(* IEC 61131-3 sources: ArdisCVDCore/codesys, 27 files *)

(* ---- E_GasChannelInit.st ---- *)
TYPE E_GasChannelInit :
(
    INIT_START,
    INIT_RAMPTIME_HOLD,
    INIT_RAMPSTEP_HOLD,
    INIT_RAMPEN_HOLD,
    INIT_MODE_HOLD,
    INIT_DONE,
    CLOSE_HOLD,
    CLOSED
);
END_TYPE

(* ---- E_MicrowaveState.st ---- *)
TYPE E_MicrowaveState :
(
    MW_IDLE,
    MW_PREHEAT_START_HOLD,
    MW_PREHEATING,
    MW_PREHEAT_READY,
    MW_RUN_START_HOLD,
    MW_RUNNING,
    MW_RUN_STOP_HOLD,
    MW_PREHEAT_ABORT_HOLD,
    MW_FAULT_STOP_HOLD,
    MW_FAULT_LATCHED
);
END_TYPE

(* ---- ST_GasChannelState.st ---- *)
TYPE ST_GasChannelState :
STRUCT
    eInit            : E_GasChannelInit;
    iInitDelay       : INT;
    xRegulating      : BOOL;
    xFaultActive     : BOOL;
    xCloseConfirmed  : BOOL;
    iLastSetpointRaw : INT;
END_STRUCT
END_TYPE

(* ---- ST_MicrowaveState.st ---- *)
TYPE ST_MicrowaveState :
STRUCT
    xLastPreheatValue    : BOOL;
    xLastOnValue         : BOOL;
    xLastResetRequest    : BOOL;
    iLastSetpointRaw     : INT;
    wFaultReason         : WORD;
    iResetHoldScans      : INT;
    iPreheatElapsedScans : INT;
END_STRUCT
END_TYPE

(* ---- GVL_Alarms.st ---- *)
VAR_GLOBAL RETAIN
    wRetainMagic      : WORD;
    wParamAlarmEnable : WORD;
    wParamAbortEnable : WORD;
    abParamAlarmPct   : ARRAY[0..6] OF BYTE;
    abParamAbortPct   : ARRAY[0..6] OF BYTE;
    wMwReflAlarmWatt  : WORD;
    wMwReflAbortWatt  : WORD;
    wTempEnable       : WORD;
    wSampleTargetC    : WORD;
    bSampleAlarmPct   : BYTE;
    abWaterTargetC    : ARRAY[0..3] OF BYTE;
    abWaterAlarmPct   : ARRAY[0..3] OF BYTE;
    abWaterAbortPct   : ARRAY[0..3] OF BYTE;
    wInputEnable      : WORD;
    wInputReaction    : WORD;
    uiLidInput        : UINT;
END_VAR

VAR_GLOBAL
    awAlarmMask     : ARRAY[0..3] OF WORD;
    awAbortMask     : ARRAY[0..3] OF WORD;
    awAbortLatched  : ARRAY[0..3] OF WORD;
    xAbortActive    : BOOL;
    xRunActive      : BOOL;
    wGpvInhibit     : WORD;
    wVpvInhibit     : WORD;
    xForeVacInhibit : BOOL;
    xTurboInhibit   : BOOL;
    xMwInhibit      : BOOL;
    xMwTripActive   : BOOL;
    wMwTripLatched  : WORD;
    xThresholdsOk   : BOOL;
    xRetainWasBlank : BOOL;
    uiAbortCount    : UINT;
END_VAR

(* ---- GVL_CoolingIO.st ---- *)
VAR_GLOBAL
    awCoolMod1Value  : ARRAY[0..7] OF WORD;
    awCoolMod1Status : ARRAY[0..7] OF WORD;

    awCoolMod2Value  : ARRAY[0..7] OF WORD;
    awCoolMod2Status : ARRAY[0..7] OF WORD;
END_VAR

(* ---- GVL_Debug.st ---- *)
VAR_GLOBAL
    uiDbgGasReinitCount : UINT;
    xDbgReboot          : BOOL;
END_VAR

(* ---- GVL_GasIO.st ---- *)
VAR_GLOBAL
    awMeasuredRaw     : ARRAY[0..5] OF WORD;
    awSetpointRaw     : ARRAY[0..5] OF WORD;
    axSetpointTrigger : ARRAY[0..5] OF BOOL;

    awModeValue       : ARRAY[0..5] OF WORD;
    axModeTrigger     : ARRAY[0..5] OF BOOL;

    awRampTimeValue   : ARRAY[0..5] OF WORD;
    axRampTimeTrigger : ARRAY[0..5] OF BOOL;

    awRampStepValue   : ARRAY[0..5] OF WORD;
    axRampStepTrigger : ARRAY[0..5] OF BOOL;

    awRampEnValue     : ARRAY[0..5] OF WORD;
    axRampEnTrigger   : ARRAY[0..5] OF BOOL;
END_VAR

(* ---- GVL_GasValveIO.st ---- *)
VAR_GLOBAL
    axGpvOutput : ARRAY[1..8] OF BOOL;
END_VAR

(* ---- GVL_MicrowaveIO.st ---- *)
VAR_GLOBAL
    awMwPowerRaw       : ARRAY[0..1] OF WORD;
    axMwStatusBlock1   : ARRAY[0..1] OF BOOL;
    axMwStatusBlock2   : ARRAY[0..5] OF BOOL;
    axMwStatusBlock3   : ARRAY[0..7] OF BOOL;

    xMwPreheatValue    : BOOL;
    xMwPreheatTrigger  : BOOL;
    xMwOnValue         : BOOL;
    xMwOnTrigger       : BOOL;
    xMwResetTrigger    : BOOL;
    wMwSetpointRaw     : WORD;
    xMwSetpointTrigger : BOOL;
END_VAR

(* ---- GVL_ModbusHolding.st ---- *)
VAR_GLOBAL
    awHolding AT %QW0 : ARRAY[0..295] OF WORD;
END_VAR

(* ---- GVL_PlcIO.st ---- *)
VAR_GLOBAL
    axFastDigitalIn : ARRAY[1..8] OF BOOL;
    axDigitalIn     : ARRAY[9..12] OF BOOL;
END_VAR

(* ---- GVL_PyroIO.st ---- *)
VAR_GLOBAL
    awPyroRxtCh1Raw     : ARRAY[0..1] OF WORD;
    awPyroRxtCh2Raw     : ARRAY[0..1] OF WORD;
    awPyroRxtRatioRaw   : ARRAY[0..1] OF WORD;
    wPyroRxtAdcStatus   : WORD;
    wPyroRxtDevStatus   : WORD;

    awPyroSmartCh1Raw   : ARRAY[0..1] OF WORD;
    awPyroSmartCh2Raw   : ARRAY[0..1] OF WORD;
    awPyroSmartRatioRaw : ARRAY[0..1] OF WORD;
    wPyroSmartAdcStatus : WORD;
    wPyroSmartDevStatus : WORD;
END_VAR

(* ---- GVL_TurboPumpIO.st ---- *)
VAR_GLOBAL
    awTurboStatusRaw  : ARRAY[0..3] OF WORD;
    wTurboTempRaw     : WORD;

    wTurboCommandValue   : WORD;
    xTurboCommandTrigger : BOOL;
END_VAR

(* ---- GVL_VacuumIO.st ---- *)
VAR_GLOBAL
    axVpvOutput : ARRAY[1..8] OF BOOL;
    xWaterPumpOutput : BOOL;
    xForeVacPumpOutput : BOOL;
END_VAR

(* ---- FB_IncrementalPid.st ---- *)
FUNCTION_BLOCK FB_IncrementalPid
VAR_INPUT
    xEnable       : BOOL;
    xReset        : BOOL;
    xDirectMode   : BOOL;
    rSetpoint     : REAL;
    rMeasured     : REAL;
    rKp           : REAL;
    rKi           : REAL;
    rKd           : REAL;
    xSmartMode    : BOOL;
    rSmartKp      : REAL;
    wPresetId     : WORD;
    rPresetOutput : REAL;
    wShiftId      : WORD;
    rShiftDelta   : REAL;
    rLowerLimit   : REAL;
    rUpperLimit   : REAL;
    rDirectValue  : REAL;
    rCycleSeconds : REAL := 0.2;
END_VAR
VAR_OUTPUT
    rError  : REAL;
    rP      : REAL;
    rI      : REAL;
    rD      : REAL;
    rOutput : REAL;
    wPresetDoneId : WORD;
    wShiftDoneId  : WORD;
END_VAR
VAR
    rPreviousError : REAL;
    xInitialized   : BOOL;
    rMin           : REAL;
    rMax           : REAL;
	arErrorBuffer      : ARRAY[0..99] OF REAL;
    i                  : INT;
    rErrAverageFirst   : REAL;
    rErrAverageLast    : REAL;
    rErrAverageIntegral : REAL;
    rKpActive           : REAL;
    wPresetSeenId       : WORD;
    xPresetArmed        : BOOL;
    rPresetFromError    : REAL;
    wShiftSeenId        : WORD;
    xShiftNew           : BOOL;
    rPresetShift        : REAL;
END_VAR

IF rLowerLimit <= rUpperLimit THEN
    rMin := rLowerLimit;
    rMax := rUpperLimit;
ELSE
    rMin := rUpperLimit;
    rMax := rLowerLimit;
END_IF;

rError := rMeasured - rSetpoint;

xShiftNew := FALSE;
IF wShiftId <> wShiftSeenId THEN
    wShiftSeenId := wShiftId;
    IF wShiftId <> WORD#0 THEN
        xShiftNew := TRUE;
        wShiftDoneId := wShiftId;
    END_IF;
END_IF;

IF NOT xEnable THEN
    rP := 0.0;
    rI := 0.0;
    rD := 0.0;
    rOutput := rMin;
    rPreviousError := rError;
    xInitialized := FALSE;
    RETURN;
END_IF;

IF xReset OR NOT xInitialized THEN
    rPreviousError := rError;
    rOutput := rMin;

    FOR i := 0 TO 99 DO
        arErrorBuffer[i] := rError;
    END_FOR;

    xInitialized := TRUE;
END_IF;

IF xShiftNew THEN
    IF xPresetArmed THEN
        rPresetShift := rPresetShift + rShiftDelta;
    ELSIF NOT xDirectMode THEN
        rOutput := rOutput + rShiftDelta;
    END_IF;
END_IF;

IF wPresetId <> wPresetSeenId THEN
    wPresetSeenId := wPresetId;
    xPresetArmed := wPresetId <> WORD#0;
    rPresetFromError := rError;
    rPresetShift := 0.0;
END_IF;

IF rCycleSeconds > 0.001 THEN
    FOR i := 0 TO 98 DO
        arErrorBuffer[i] := arErrorBuffer[i + 1];
    END_FOR;
    arErrorBuffer[99] := rError;

    rErrAverageFirst := 0.0;
    FOR i := 87 TO 91 DO
        rErrAverageFirst := rErrAverageFirst + arErrorBuffer[i];
    END_FOR;
    rErrAverageFirst := rErrAverageFirst / 5.0;

    rErrAverageLast := 0.0;
    FOR i := 98 TO 99 DO
        rErrAverageLast := rErrAverageLast + arErrorBuffer[i];
    END_FOR;
    rErrAverageLast := rErrAverageLast / 2.0;

    rD := rKd * (rErrAverageLast - rErrAverageFirst);

    rErrAverageIntegral := 0.0;
    FOR i := 80 TO 99 DO
        rErrAverageIntegral := rErrAverageIntegral + arErrorBuffer[i];
    END_FOR;
    rErrAverageIntegral := rErrAverageIntegral / 20.0;

    rI := rKi * rErrAverageIntegral;
ELSE
    rD := 0.0;
    rI := 0.0;
END_IF;

IF xSmartMode AND rError > 0.0 AND rD > 0.0 THEN
    rKpActive := rSmartKp;
ELSE
    rKpActive := rKp;
END_IF;

rP := rKpActive * rError;

rPreviousError := rError;

IF xDirectMode THEN
    rOutput := rDirectValue;
    rPresetFromError := rError;
ELSIF xPresetArmed AND rError * rPresetFromError <= 0.0 THEN
    rOutput := rPresetOutput + rPresetShift;
    xPresetArmed := FALSE;
    wPresetDoneId := wPresetSeenId;
ELSE
    rOutput := rOutput + rP + rI + rD;
END_IF;

IF rOutput > rMax THEN
    rOutput := rMax;
ELSIF rOutput < rMin THEN
    rOutput := rMin;
END_IF;

(* ---- FB_ThyracontAscii.st ---- *)
FUNCTION_BLOCK FB_ThyracontAscii
VAR_INPUT
    xEnable : BOOL := TRUE;
    udiPort : UDINT := 1;
    udiAddress : UDINT := 1;
    udiBaudrate : UDINT := 9600;
    tPollInterval : TIME := T#1S;
END_VAR
VAR_OUTPUT
    xValid : BOOL;
    xConnected : BOOL;
    rPressureMbar : REAL;
    rPressureTorr : REAL;
    wStatusFlags : WORD;
    wErrorCode : WORD;
    udiCycle : UDINT;
END_VAR
VAR
    fbOpen : COM.Open;
    fbWrite : COM.Write;
    fbRead : COM.Read;
    aParams : ARRAY[1..7] OF COM.PARAMETER;
    hCom : CAA.HANDLE;
    aTx : ARRAY[0..9] OF BYTE := [BYTE#48, BYTE#48, BYTE#49, BYTE#48, BYTE#77, BYTE#86, BYTE#48, BYTE#48, BYTE#68, BYTE#13];
    aRx : ARRAY[0..63] OF BYTE;
    aAdr : ARRAY[0..2] OF BYTE;
    iAddr : INT;
    iChecksum : INT;
    iState : INT;
    udiPollTicks : UDINT;
    udiPollTicksMax : UDINT := 5;
    xOpenExecute : BOOL;
    xWriteExecute : BOOL;
    xReadExecute : BOOL;
    i : INT;
    j : INT;
    iSize : INT;
    iFrameStart : INT;
    iDataLen : INT;
    iDataStart : INT;
    iDigit : INT;
    iSign : INT;
    iExpSign : INT;
    iExp : INT;
    rParsed : REAL;
    rDiv : REAL;
    xFraction : BOOL;
    xExponent : BOOL;
    xHasDigit : BOOL;
END_VAR

IF NOT xEnable THEN
    xOpenExecute := FALSE;
    xWriteExecute := FALSE;
    xReadExecute := FALSE;
    xConnected := FALSE;
    xValid := FALSE;
    wStatusFlags := WORD#0;
    wErrorCode := WORD#0;
    iState := 0;
    RETURN;
END_IF;

aParams[1].udiParameterId := COM.CAA_Parameter_Constants.udiPort;
aParams[1].udiValue := udiPort;
aParams[2].udiParameterId := COM.CAA_Parameter_Constants.udiBaudrate;
aParams[2].udiValue := udiBaudrate;
aParams[3].udiParameterId := COM.CAA_Parameter_Constants.udiParity;
aParams[3].udiValue := 2;
aParams[4].udiParameterId := COM.CAA_Parameter_Constants.udiStopBits;
aParams[4].udiValue := 0;
aParams[5].udiParameterId := COM.CAA_Parameter_Constants.udiTimeout;
aParams[5].udiValue := 200000;
aParams[6].udiParameterId := COM.CAA_Parameter_Constants.udiByteSize;
aParams[6].udiValue := 8;
aParams[7].udiParameterId := COM.CAA_Parameter_Constants.udiBinary;
aParams[7].udiValue := 1;

iAddr := UDINT_TO_INT(udiAddress);
IF (iAddr < 1) OR (iAddr > 16) THEN
    iAddr := 1;
END_IF;
aAdr[0] := INT_TO_BYTE(iAddr / 100 MOD 10 + 48);
aAdr[1] := INT_TO_BYTE(iAddr / 10 MOD 10 + 48);
aAdr[2] := INT_TO_BYTE(iAddr MOD 10 + 48);
aTx[0] := aAdr[0];
aTx[1] := aAdr[1];
aTx[2] := aAdr[2];

iChecksum := 0;
FOR i := 0 TO 7 DO
    iChecksum := iChecksum + BYTE_TO_INT(aTx[i]);
END_FOR;
aTx[8] := INT_TO_BYTE(iChecksum MOD 64 + 64);

IF tPollInterval <= T#0MS THEN
    udiPollTicksMax := 0;
ELSIF tPollInterval <= T#200MS THEN
    udiPollTicksMax := 1;
ELSE
    udiPollTicksMax := TIME_TO_UDINT(tPollInterval) / 200;
    IF udiPollTicksMax < 1 THEN
        udiPollTicksMax := 1;
    END_IF;
END_IF;

CASE iState OF
    0:
        xOpenExecute := TRUE;
        xConnected := FALSE;
        xValid := FALSE;
        wErrorCode := WORD#1;
        IF fbOpen.xDone THEN
            hCom := fbOpen.hCom;
            xOpenExecute := FALSE;
            xConnected := TRUE;
            wErrorCode := WORD#0;
            iState := 10;
        ELSIF fbOpen.xError THEN
            xOpenExecute := FALSE;
            wErrorCode := WORD#2;
            iState := 50;
        END_IF;

    10:
        udiPollTicks := 0;
        FOR i := 0 TO 63 DO
            aRx[i] := BYTE#0;
        END_FOR;
        xWriteExecute := TRUE;
        iState := 20;

    20:
        IF fbWrite.xDone THEN
            xWriteExecute := FALSE;
            xReadExecute := TRUE;
            iState := 30;
        ELSIF fbWrite.xError THEN
            xWriteExecute := FALSE;
            xValid := FALSE;
            wErrorCode := WORD#3;
            iState := 50;
        END_IF;

    30:
        IF fbRead.xDone THEN
            xReadExecute := FALSE;
            iSize := UDINT_TO_INT(fbRead.szSize);
            iFrameStart := -1;

            IF iSize >= 10 THEN
                FOR i := 0 TO iSize - 8 DO
                    IF (aRx[i] = aAdr[0]) AND (aRx[i + 1] = aAdr[1]) AND
                       (aRx[i + 2] = aAdr[2]) AND (aRx[i + 3] = BYTE#49) AND
                       (aRx[i + 4] = BYTE#77) AND (aRx[i + 5] = BYTE#86) THEN
                        iFrameStart := i;
                        EXIT;
                    END_IF;
                END_FOR;
            END_IF;

            IF iFrameStart < 0 THEN
                xValid := FALSE;
                wErrorCode := WORD#5;
                iState := 50;
            ELSE
                iDataLen := (BYTE_TO_INT(aRx[iFrameStart + 6]) - 48) * 10 +
                            (BYTE_TO_INT(aRx[iFrameStart + 7]) - 48);
                iDataStart := iFrameStart + 8;

                IF (iDataLen <= 0) OR ((iDataStart + iDataLen) >= iSize) THEN
                    xValid := FALSE;
                    wErrorCode := WORD#6;
                    iState := 50;
                ELSE
                    rParsed := 0.0;
                    rDiv := 10.0;
                    iSign := 1;
                    iExpSign := 1;
                    iExp := 0;
                    xFraction := FALSE;
                    xExponent := FALSE;
                    xHasDigit := FALSE;

                    FOR i := 0 TO iDataLen - 1 DO
                        j := iDataStart + i;
                        IF (aRx[j] >= BYTE#48) AND (aRx[j] <= BYTE#57) THEN
                            iDigit := BYTE_TO_INT(aRx[j]) - 48;
                            xHasDigit := TRUE;
                            IF xExponent THEN
                                iExp := iExp * 10 + iDigit;
                            ELSIF xFraction THEN
                                rParsed := rParsed + INT_TO_REAL(iDigit) / rDiv;
                                rDiv := rDiv * 10.0;
                            ELSE
                                rParsed := rParsed * 10.0 + INT_TO_REAL(iDigit);
                            END_IF;
                        ELSIF aRx[j] = BYTE#45 THEN
                            IF xExponent THEN
                                iExpSign := -1;
                            ELSE
                                iSign := -1;
                            END_IF;
                        ELSIF (aRx[j] = BYTE#46) OR (aRx[j] = BYTE#44) THEN
                            xFraction := TRUE;
                        ELSIF (aRx[j] = BYTE#69) OR (aRx[j] = BYTE#101) THEN
                            xExponent := TRUE;
                        END_IF;
                    END_FOR;

                    IF xHasDigit THEN
                        IF iExp > 38 THEN
                            iExp := 38;
                        END_IF;

                        FOR i := 1 TO iExp DO
                            IF iExpSign > 0 THEN
                                rParsed := rParsed * 10.0;
                            ELSE
                                rParsed := rParsed / 10.0;
                            END_IF;
                        END_FOR;

                        rPressureMbar := rParsed * INT_TO_REAL(iSign);
                        rPressureTorr := rPressureMbar * 0.7500637;
                        xValid := TRUE;
                        xConnected := TRUE;
                        wErrorCode := WORD#0;
                        udiCycle := udiCycle + 1;
                    ELSE
                        xValid := FALSE;
                        wErrorCode := WORD#7;
                    END_IF;

                    iState := 50;
                END_IF;
            END_IF;
        ELSIF fbRead.xError THEN
            xReadExecute := FALSE;
            xValid := FALSE;
            wErrorCode := WORD#4;
            iState := 50;
        END_IF;

    50:
        udiPollTicks := udiPollTicks + 1;
        IF udiPollTicks >= udiPollTicksMax THEN
            iState := 10;
        END_IF;

ELSE
    iState := 0;
END_CASE;

wStatusFlags := WORD#0;
IF xValid THEN
    wStatusFlags := wStatusFlags OR WORD#16#0001;
END_IF;

fbOpen(
    xExecute := xOpenExecute,
    usiListLength := 7,
    pParameterList := ADR(aParams));

fbWrite(
    xExecute := xWriteExecute,
    udiTimeOut := 100000,
    hCom := hCom,
    pBuffer := ADR(aTx),
    szSize := SIZEOF(aTx));

fbRead(
    xExecute := xReadExecute,
    udiTimeOut := 300000,
    hCom := hCom,
    pBuffer := ADR(aRx),
    szBuffer := SIZEOF(aRx));

(* ---- PLC_PRG.st ---- *)
PROGRAM PLC_PRG
(* main program: hmi link, signal tower, pressure pid *)
VAR
    xDoBlinkTest : BOOL;
    wBenchMuAo1Output : ARRAY[0..0] OF WORD;
    xTrafficLightGreen  : BOOL;
    xTrafficLightYellow : BOOL;
    xTrafficLightRed    : BOOL;
    wTrafficLightMask   : WORD;

    xHmiWriteSeen         : BOOL;
    udiHmiStaleCycles     : UDINT;
    xHmiLinkLost          : BOOL;

    awMvAi1Value  : ARRAY[0..1] OF WORD;
    awMvAi1Status : ARRAY[0..0] OF WORD;
    uMvAi1Value   : U_DWORD_REAL;
    wMvAi1Status  : WORD;
    xMvAi1Ok      : BOOL;
    rMvAi1Percent : REAL;
    rMvAi1Voltage : REAL;
    rChMeasuredMv : REAL;

	wDiscreteInputs : WORD;
    iDiIndex        : INT;

    rChamberMuAo1Command : REAL;
    xChamberMuAo1Clamped : BOOL;
    uiChamberMuAo1Command : UINT;
    fbChamber : FB_IncrementalPid;
    fbPlenum  : FB_IncrementalPid;
    xProtocolOk    : BOOL;
    xChamberEnable : BOOL;
    xPlenumEnable  : BOOL;
    xReset         : BOOL;
    udiCycle       : UDINT;
    rChSetpoint : REAL;
    rChMeasured : REAL;
    rChKp       : REAL;
    rChKi       : REAL;
    rChKd       : REAL;
    rChLower    : REAL;
    rChUpper    : REAL;
    rChDirect   : REAL;
    rChSmartKp  : REAL;
    xChSmartMode : BOOL;
    rChPresetOutput : REAL;
    wChPresetId     : WORD;
    rChShiftDelta   : REAL;
    wChShiftId      : WORD;
    rPlSetpoint : REAL;
    rPlMeasured : REAL;
    rPlKp       : REAL;
    rPlKi       : REAL;
    rPlKd       : REAL;
    rPlLower    : REAL;
    rPlUpper    : REAL;
    rPlDirect   : REAL;
    dwValue     : DWORD;
    xDoBlinkTestEnable : BOOL;
    xBenchMuAo1Enable : BOOL;
    xBenchMuAo1Clamped : BOOL;
    uiBenchMuAo1Command : UINT;
    uiBenchMuAo1Applied : UINT;
    awMvAi1Raw : ARRAY[0..1] OF WORD;
END_VAR
VAR CONSTANT
    HMI_STALE_CYCLES  : UDINT := UDINT#15;
END_VAR

(* commands from the hmi *)
xProtocolOk := awHolding[0] = WORD#1;
xChamberEnable := xProtocolOk AND (awHolding[1] AND WORD#16#0001) <> WORD#0;
xPlenumEnable := xProtocolOk AND (awHolding[1] AND WORD#16#0002) <> WORD#0;
xReset := (awHolding[1] AND WORD#16#0004) <> WORD#0;
xTrafficLightGreen  := (awHolding[1] AND WORD#16#0010) <> WORD#0;
xTrafficLightYellow := (awHolding[1] AND WORD#16#0020) <> WORD#0;
xTrafficLightRed    := (awHolding[1] AND WORD#16#0040) <> WORD#0;

(* hmi watchdog: link lost after 3 s without a write *)
xHmiWriteSeen := (awHolding[1] AND WORD#16#8000) = WORD#0;

IF xHmiWriteSeen THEN
    udiHmiStaleCycles := UDINT#0;
ELSIF udiHmiStaleCycles < HMI_STALE_CYCLES THEN
    udiHmiStaleCycles := udiHmiStaleCycles + UDINT#1;
END_IF;

xHmiLinkLost := udiHmiStaleCycles >= HMI_STALE_CYCLES;

(* signal tower, all three lamps on when the link is lost *)
wTrafficLightMask := WORD#0;
IF xHmiLinkLost THEN
    wTrafficLightMask := WORD#16#0007;
ELSE
    IF xTrafficLightGreen THEN
        wTrafficLightMask := wTrafficLightMask OR WORD#16#0001;
    END_IF;
    IF xTrafficLightYellow THEN
        wTrafficLightMask := wTrafficLightMask OR WORD#16#0002;
    END_IF;
    IF xTrafficLightRed THEN
        wTrafficLightMask := wTrafficLightMask OR WORD#16#0004;
    END_IF;
END_IF;

(* set the marker, the hmi clears it on its next write *)
awHolding[1] := awHolding[1] OR WORD#16#8000;

(* chamber pid output to the analogue output, max 500 *)
rChamberMuAo1Command := fbChamber.rOutput / 10.0;
xChamberMuAo1Clamped := rChamberMuAo1Command > 500.0;

IF xChamberMuAo1Clamped THEN
    uiChamberMuAo1Command := UINT#500;
ELSE
    uiChamberMuAo1Command := REAL_TO_UINT(rChamberMuAo1Command);
END_IF;

(* chamber pressure from the analogue input module *)
wMvAi1Status := awMvAi1Status[0];
xMvAi1Ok := wMvAi1Status = WORD#16#0000;

uMvAi1Value.dwValue := SHL(WORD_TO_DWORD(awMvAi1Value[1]), 16) OR WORD_TO_DWORD(awMvAi1Value[0]);
rMvAi1Percent := uMvAi1Value.rValue;
rMvAi1Voltage := LIMIT(0.0, rMvAi1Percent / 10.0, 10.0);

IF xMvAi1Ok THEN
    rChMeasuredMv := LIMIT(0.0, rMvAi1Percent * 10.0, 1000.0);
END_IF;

(* pid setpoints and gains from the hmi *)
rChSetpoint := F_ReadFixed(awHolding[4], awHolding[5]);
rChMeasured := rChMeasuredMv;
rChKp := F_ReadFixed(awHolding[8], awHolding[9]);
rChKi := F_ReadFixed(awHolding[10], awHolding[11]);
rChKd := F_ReadFixed(awHolding[12], awHolding[13]);
rChLower := F_ReadFixed(awHolding[14], awHolding[15]);
rChUpper := F_ReadFixed(awHolding[16], awHolding[17]);
rChDirect := F_ReadFixed(awHolding[18], awHolding[19]);
rChSmartKp := F_ReadFixed(awHolding[27], awHolding[28]);
xChSmartMode := awHolding[29] <> WORD#0;
rChPresetOutput := F_ReadFixed(awHolding[56], awHolding[57]);
wChPresetId := awHolding[58];
rChShiftDelta := F_ReadFixed(awHolding[59], awHolding[60]);
wChShiftId := awHolding[61];

rPlSetpoint := F_ReadFixed(awHolding[30], awHolding[31]);
rPlMeasured := F_ReadFixed(awHolding[32], awHolding[33]);
rPlKp := F_ReadFixed(awHolding[34], awHolding[35]);
rPlKi := F_ReadFixed(awHolding[36], awHolding[37]);
rPlKd := F_ReadFixed(awHolding[38], awHolding[39]);
rPlLower := F_ReadFixed(awHolding[40], awHolding[41]);
rPlUpper := F_ReadFixed(awHolding[42], awHolding[43]);
rPlDirect := F_ReadFixed(awHolding[44], awHolding[45]);

(* chamber pid *)
fbChamber(
    xEnable := xChamberEnable,
    xReset := xReset,
    xDirectMode := awHolding[20] <> WORD#0,
    rSetpoint := rChSetpoint,
    rMeasured := rChMeasured,
    rKp := rChKp,
    rKi := rChKi,
    rKd := rChKd,
    xSmartMode := xChSmartMode,
    rSmartKp := rChSmartKp,
    wPresetId := wChPresetId,
    rPresetOutput := rChPresetOutput,
    wShiftId := wChShiftId,
    rShiftDelta := rChShiftDelta,
    rLowerLimit := rChLower,
    rUpperLimit := rChUpper,
    rDirectValue := rChDirect,
    rCycleSeconds := 0.2);

(* plenum pid *)
fbPlenum(
    xEnable := xPlenumEnable,
    xReset := xReset,
    xDirectMode := awHolding[46] <> WORD#0,
    rSetpoint := rPlSetpoint,
    rMeasured := rPlMeasured,
    rKp := rPlKp,
    rKi := rPlKi,
    rKd := rPlKd,
    rLowerLimit := rPlLower,
    rUpperLimit := rPlUpper,
    rDirectValue := rPlDirect,
    rCycleSeconds := 0.2);

(* cycle counter and blink test *)
udiCycle := udiCycle + 1;
xDoBlinkTestEnable := awHolding[150] = WORD#16#A55A;
xDoBlinkTest := xDoBlinkTestEnable AND ((udiCycle MOD UDINT#10) < UDINT#5);

(* to the hmi: version, status, cycle counter *)
awHolding[100] := WORD#1;
IF xProtocolOk THEN
    awHolding[101] := WORD#16#0003;
ELSE
    awHolding[101] := WORD#0;
END_IF;
awHolding[102] := DWORD_TO_WORD(udiCycle);
awHolding[103] := DWORD_TO_WORD(SHR(udiCycle, 16));

(* chamber pid terms to the hmi *)
dwValue := F_ToFixed(fbChamber.rError);
awHolding[104] := DWORD_TO_WORD(dwValue);
awHolding[105] := DWORD_TO_WORD(SHR(dwValue, 16));
dwValue := F_ToFixed(fbChamber.rP);
awHolding[106] := DWORD_TO_WORD(dwValue);
awHolding[107] := DWORD_TO_WORD(SHR(dwValue, 16));
dwValue := F_ToFixed(fbChamber.rI);
awHolding[108] := DWORD_TO_WORD(dwValue);
awHolding[109] := DWORD_TO_WORD(SHR(dwValue, 16));
dwValue := F_ToFixed(fbChamber.rD);
awHolding[110] := DWORD_TO_WORD(dwValue);
awHolding[111] := DWORD_TO_WORD(SHR(dwValue, 16));
dwValue := F_ToFixed(fbChamber.rOutput);
awHolding[112] := DWORD_TO_WORD(dwValue);
awHolding[113] := DWORD_TO_WORD(SHR(dwValue, 16));
awHolding[114] := fbChamber.wPresetDoneId;
awHolding[115] := fbChamber.wShiftDoneId;

(* plenum pid terms to the hmi *)
dwValue := F_ToFixed(fbPlenum.rError);
awHolding[120] := DWORD_TO_WORD(dwValue);
awHolding[121] := DWORD_TO_WORD(SHR(dwValue, 16));
dwValue := F_ToFixed(fbPlenum.rP);
awHolding[122] := DWORD_TO_WORD(dwValue);
awHolding[123] := DWORD_TO_WORD(SHR(dwValue, 16));
dwValue := F_ToFixed(fbPlenum.rI);
awHolding[124] := DWORD_TO_WORD(dwValue);
awHolding[125] := DWORD_TO_WORD(SHR(dwValue, 16));
dwValue := F_ToFixed(fbPlenum.rD);
awHolding[126] := DWORD_TO_WORD(dwValue);
awHolding[127] := DWORD_TO_WORD(SHR(dwValue, 16));
dwValue := F_ToFixed(fbPlenum.rOutput);
awHolding[128] := DWORD_TO_WORD(dwValue);
awHolding[129] := DWORD_TO_WORD(SHR(dwValue, 16));

(* chamber pressure and sensor status to the hmi *)
dwValue := F_ToFixed(rChMeasuredMv);
awHolding[130] := DWORD_TO_WORD(dwValue);
awHolding[131] := DWORD_TO_WORD(SHR(dwValue, 16));
awHolding[132] := wMvAi1Status;

(* discrete inputs to the hmi *)
wDiscreteInputs := WORD#0;
FOR iDiIndex := 1 TO 8 DO
    IF axFastDigitalIn[iDiIndex] THEN
        wDiscreteInputs := wDiscreteInputs OR SHL(WORD#1, iDiIndex - 1);
    END_IF;
END_FOR;
FOR iDiIndex := 9 TO 12 DO
    IF axDigitalIn[iDiIndex] THEN
        wDiscreteInputs := wDiscreteInputs OR SHL(WORD#1, iDiIndex - 1);
    END_IF;
END_FOR;
awHolding[139] := wDiscreteInputs;

(* manual analogue output test from the hmi *)
uiBenchMuAo1Command := WORD_TO_UINT(awHolding[154]);
xBenchMuAo1Enable := awHolding[155] = WORD#16#A55A;
xBenchMuAo1Clamped := uiBenchMuAo1Command > UINT#500;

IF xBenchMuAo1Clamped THEN
    uiBenchMuAo1Command := UINT#500;
END_IF;

IF xBenchMuAo1Enable THEN
    uiBenchMuAo1Applied := uiBenchMuAo1Command;
ELSE
    uiBenchMuAo1Applied := UINT#0;
END_IF;

(* test flags to the hmi *)
IF xBenchMuAo1Enable THEN
    awHolding[157] := awHolding[157] OR WORD#16#0001;
END_IF;

IF xBenchMuAo1Clamped THEN
    awHolding[157] := awHolding[157] OR WORD#16#0002;
END_IF;

(* output command from the chamber pid *)
IF fbChamber.rOutput <= 0.0 THEN
    uiChamberMuAo1Command := UINT#0;
    xChamberMuAo1Clamped := FALSE;
ELSE
    rChamberMuAo1Command := fbChamber.rOutput / 10.0;
    xChamberMuAo1Clamped := rChamberMuAo1Command > 500.0;

    IF xChamberMuAo1Clamped THEN
        uiChamberMuAo1Command := UINT#500;
    ELSE
        uiChamberMuAo1Command := REAL_TO_UINT(rChamberMuAo1Command);
    END_IF;
END_IF;

(* drive the output: test value, pid or zero *)
IF xBenchMuAo1Enable THEN
    uiBenchMuAo1Applied := uiBenchMuAo1Command;
ELSIF xChamberEnable THEN
    uiBenchMuAo1Applied := uiChamberMuAo1Command;
ELSE
    uiBenchMuAo1Applied := UINT#0;
END_IF;

wBenchMuAo1Output[0] := UINT_TO_WORD(uiBenchMuAo1Applied);
awHolding[156] := wBenchMuAo1Output[0];

(* ---- PRG_Alarms.st ---- *)
PROGRAM PRG_Alarms
(* alarms and abort *)
VAR
    i : INT;
    iBase : INT;
    iBit : INT;
    iWord : INT;

    xFirstScan : BOOL := TRUE;

    axAlarm : ARRAY[0..63] OF BOOL;
    axAbort : ARRAY[0..63] OF BOOL;

    arBandSetpoint : ARRAY[0..6] OF REAL;
    arBandMeasured : ARRAY[0..6] OF REAL;
    axBandGate     : ARRAY[0..6] OF BOOL;

    arWaterTempC : ARRAY[0..3] OF REAL;
    axWaterTempValid : ARRAY[0..3] OF BOOL;

    rSetpoint : REAL;
    rMeasured : REAL;
    rBand     : REAL;
    rReflKw   : REAL;
    rSampleC  : REAL;
    rFlowLpm  : REAL;
    rWaterBar : REAL;
    rCdaBar   : REAL;

    wCommand    : WORD;
    wStatusWord : WORD;
    wMwStatus : WORD;
    wTempValid : WORD;
    wFlowValid : WORD;
    wTurboStatus : WORD;
    wDiscrete : WORD;
    wMwTripNow : WORD;

    xMwRequested : BOOL;
    xPyroValid : BOOL;
    xTurboAnswering : BOOL;
    xWaterPump : BOOL;
    xFlowArmed : BOOL;
    xLidClosed : BOOL;

    xAnyAlarm : BOOL;
    xAnyAbort : BOOL;

    xReset : BOOL;
    xResetPrev : BOOL;

    fbFlowArm : TON;
END_VAR
VAR CONSTANT
    C_BLOCK_MAGIC  : WORD := WORD#16#A500;
    C_RETAIN_MAGIC : WORD := WORD#16#5A5A;

    C_FLOW_MIN_LOW  : REAL := 1.0;
    C_FLOW_MIN_HIGH : REAL := 5.0;

    C_WATER_ALARM_BAR : REAL := 0.7;
    C_WATER_ABORT_BAR : REAL := 0.5;
    C_CDA_ALARM_BAR   : REAL := 5.0;
    C_CDA_ABORT_BAR   : REAL := 4.0;

    C_CHAMBER_MAX_TORR : REAL := 800.0;
    C_HMI_PROTOCOL     : WORD := WORD#16#0200;
    C_FLOW_ARM_TIME    : TIME := T#4S;

    C_CIRC_STAGE    : INT := 0;
    C_CIRC_CHAMBER  : INT := 1;
    C_CIRC_MWHEAD   : INT := 2;
    C_CIRC_MWPOWER  : INT := 3;
    C_CIRC_INTERNAL : INT := 5;
    C_CIRC_EXTERNAL : INT := 6;
END_VAR

(* first scan: all alarms off if the retain memory was lost *)
IF xFirstScan THEN
    xFirstScan := FALSE;
    IF wRetainMagic <> C_RETAIN_MAGIC THEN
        xRetainWasBlank := TRUE;
        wRetainMagic := C_RETAIN_MAGIC;
        wParamAlarmEnable := WORD#0;
        wParamAbortEnable := WORD#0;
        wTempEnable := WORD#0;
        wInputEnable := WORD#0;
        uiLidInput := UINT#1;
    ELSE
        xRetainWasBlank := FALSE;
    END_IF;
END_IF;

(* alarm thresholds from the hmi *)
xThresholdsOk := (awHolding[248] AND WORD#16#FF00) = C_BLOCK_MAGIC;

IF xThresholdsOk THEN
    wParamAlarmEnable := awHolding[249];
    wParamAbortEnable := awHolding[250];
    FOR i := 0 TO 6 DO
        abParamAlarmPct[i] := WORD_TO_BYTE(awHolding[251 + i] AND WORD#16#00FF);
        abParamAbortPct[i] := WORD_TO_BYTE(SHR(awHolding[251 + i], 8));
    END_FOR;
    wMwReflAlarmWatt := awHolding[258];
    wMwReflAbortWatt := awHolding[259];

    wTempEnable := awHolding[260];
    wSampleTargetC := awHolding[261];
    bSampleAlarmPct := WORD_TO_BYTE(awHolding[262] AND WORD#16#00FF);
    abWaterTargetC[0] := WORD_TO_BYTE(awHolding[263] AND WORD#16#00FF);
    abWaterTargetC[1] := WORD_TO_BYTE(SHR(awHolding[263], 8));
    abWaterTargetC[2] := WORD_TO_BYTE(awHolding[264] AND WORD#16#00FF);
    abWaterTargetC[3] := WORD_TO_BYTE(SHR(awHolding[264], 8));
    FOR i := 0 TO 3 DO
        abWaterAlarmPct[i] := WORD_TO_BYTE(awHolding[265 + i] AND WORD#16#00FF);
        abWaterAbortPct[i] := WORD_TO_BYTE(SHR(awHolding[265 + i], 8));
    END_FOR;

    wInputEnable := awHolding[269];
    wInputReaction := awHolding[270];
    xRunActive := (awHolding[271] AND WORD#16#0001) <> WORD#0;
    uiLidInput := WORD_TO_UINT(SHR(awHolding[271], 8));
    IF (uiLidInput < UINT#1) OR (uiLidInput > UINT#12) THEN
        uiLidInput := UINT#1;
    END_IF;
ELSE
    xRunActive := FALSE;
END_IF;

(* rebuild every alarm from scratch each cycle *)
FOR i := 0 TO 63 DO
    axAlarm[i] := FALSE;
    axAbort[i] := FALSE;
END_FOR;

(* inputs from the register map *)
wMwStatus := awHolding[195];
wCommand := awHolding[192];
xMwRequested := ((wCommand AND WORD#16#0003) <> WORD#0) AND (NOT xAbortActive) AND (NOT xMwInhibit)
    AND (NOT xMwTripActive);
rReflKw := F_ReadFixed(awHolding[199], awHolding[200]);

wTempValid := awHolding[238];
wFlowValid := awHolding[239];
wTurboStatus := awHolding[245];
xTurboAnswering := (awHolding[247] AND WORD#16#0001) <> WORD#0;
wDiscrete := awHolding[139];
xLidClosed := (wDiscrete AND SHL(WORD#1, UINT_TO_INT(uiLidInput) - 1)) <> WORD#0;

xWaterPump := xWaterPumpOutput;
fbFlowArm(IN := xWaterPump, PT := C_FLOW_ARM_TIME);
xFlowArmed := fbFlowArm.Q;

xPyroValid := (awHolding[166] AND WORD#16#0001) <> WORD#0;

(* chamber pressure and gases: setpoint, measured value, when to check *)
arBandSetpoint[0] := F_ReadFixed(awHolding[4], awHolding[5]);
arBandMeasured[0] := F_ReadFixed(awHolding[130], awHolding[131]);
axBandGate[0] := TRUE;

FOR i := 0 TO 5 DO
    iBase := 66 + i*5;
    arBandSetpoint[i + 1] := F_ReadFixed(awHolding[iBase], awHolding[iBase + 1]);
    arBandMeasured[i + 1] := F_ReadFixed(awHolding[iBase + 2], awHolding[iBase + 3]);
    axBandGate[i + 1] := axGpvOutput[i + 1] AND axGpvOutput[8]
        AND ((awHolding[96] AND SHL(WORD#1, i)) = WORD#0);
END_FOR;

(* deviation from the setpoint beyond the band *)
FOR i := 0 TO 6 DO
    rSetpoint := arBandSetpoint[i];
    rMeasured := arBandMeasured[i];

    IF axBandGate[i] AND (rSetpoint > 0.0) THEN
        IF (wParamAlarmEnable AND SHL(WORD#1, i)) <> WORD#0 THEN
            rBand := rSetpoint * BYTE_TO_REAL(abParamAlarmPct[i]) / 100.0;
            IF (rMeasured >= rSetpoint + rBand) OR (rMeasured <= rSetpoint - rBand) THEN
                axAlarm[i] := TRUE;
            END_IF;
        END_IF;
        IF (wParamAbortEnable AND SHL(WORD#1, i)) <> WORD#0 THEN
            rBand := rSetpoint * BYTE_TO_REAL(abParamAbortPct[i]) / 100.0;
            IF (rMeasured >= rSetpoint + rBand) OR (rMeasured <= rSetpoint - rBand) THEN
                axAbort[i] := TRUE;
            END_IF;
        END_IF;
    END_IF;
END_FOR;

(* reflected microwave power *)
IF (wParamAlarmEnable AND WORD#16#0080) <> WORD#0 THEN
    IF rReflKw * 1000.0 >= UINT_TO_REAL(WORD_TO_UINT(wMwReflAlarmWatt)) THEN
        axAlarm[7] := TRUE;
    END_IF;
END_IF;
IF (wParamAbortEnable AND WORD#16#0080) <> WORD#0 THEN
    IF rReflKw * 1000.0 >= UINT_TO_REAL(WORD_TO_UINT(wMwReflAbortWatt)) THEN
        axAbort[7] := TRUE;
    END_IF;
END_IF;

(* sample temperature from the pyrometer *)
rSampleC := F_ReadFixed(awHolding[160], awHolding[161]);
IF xPyroValid AND ((wTempEnable AND WORD#16#0001) <> WORD#0)
    AND (wSampleTargetC > WORD#0) THEN
    rSetpoint := UINT_TO_REAL(WORD_TO_UINT(wSampleTargetC));
    rBand := rSetpoint * BYTE_TO_REAL(bSampleAlarmPct) / 100.0;
    IF (rSampleC >= rSetpoint + rBand) OR (rSampleC <= rSetpoint - rBand) THEN
        axAlarm[8] := TRUE;
    END_IF;
END_IF;

(* cooling water temperatures, only while the water pump runs *)
arWaterTempC[0] := F_ReadFixed(awHolding[206 + 2*C_CIRC_INTERNAL], awHolding[207 + 2*C_CIRC_INTERNAL]);
arWaterTempC[1] := F_ReadFixed(awHolding[206 + 2*C_CIRC_EXTERNAL], awHolding[207 + 2*C_CIRC_EXTERNAL]);
arWaterTempC[2] := F_ReadFixed(awHolding[206 + 2*C_CIRC_STAGE], awHolding[207 + 2*C_CIRC_STAGE]);
arWaterTempC[3] := F_ReadFixed(awHolding[206 + 2*C_CIRC_CHAMBER], awHolding[207 + 2*C_CIRC_CHAMBER]);

axWaterTempValid[0] := (wTempValid AND SHL(WORD#1, C_CIRC_INTERNAL)) <> WORD#0;
axWaterTempValid[1] := (wTempValid AND SHL(WORD#1, C_CIRC_EXTERNAL)) <> WORD#0;
axWaterTempValid[2] := (wTempValid AND SHL(WORD#1, C_CIRC_STAGE)) <> WORD#0;
axWaterTempValid[3] := (wTempValid AND SHL(WORD#1, C_CIRC_CHAMBER)) <> WORD#0;

FOR i := 0 TO 3 DO
    IF xWaterPump AND axWaterTempValid[i] AND (abWaterTargetC[i] > BYTE#0) THEN
        rSetpoint := BYTE_TO_REAL(abWaterTargetC[i]);
        rMeasured := arWaterTempC[i];
        IF (wTempEnable AND SHL(WORD#1, i + 1)) <> WORD#0 THEN
            rBand := rSetpoint * BYTE_TO_REAL(abWaterAlarmPct[i]) / 100.0;
            IF (rMeasured >= rSetpoint + rBand) OR (rMeasured <= rSetpoint - rBand) THEN
                axAlarm[9 + i] := TRUE;
            END_IF;
        END_IF;
        IF (wTempEnable AND SHL(WORD#1, i + 9)) <> WORD#0 THEN
            rBand := rSetpoint * BYTE_TO_REAL(abWaterAbortPct[i]) / 100.0;
            IF (rMeasured >= rSetpoint + rBand) OR (rMeasured <= rSetpoint - rBand) THEN
                axAbort[9 + i] := TRUE;
            END_IF;
        END_IF;
    END_IF;
END_FOR;

(* cooling water flows, armed 4 s after the pump starts *)
FOR i := 0 TO 5 DO
    CASE i OF
        0: iBase := C_CIRC_STAGE;
        1: iBase := C_CIRC_CHAMBER;
        2: iBase := C_CIRC_MWHEAD;
        3: iBase := C_CIRC_MWPOWER;
        4: iBase := C_CIRC_INTERNAL;
    ELSE
        iBase := C_CIRC_EXTERNAL;
    END_CASE;

    IF i < 4 THEN
        rSetpoint := C_FLOW_MIN_LOW;
    ELSE
        rSetpoint := C_FLOW_MIN_HIGH;
    END_IF;

    rFlowLpm := F_ReadFixed(awHolding[220 + 2*iBase], awHolding[221 + 2*iBase]);

    IF xWaterPump AND xFlowArmed
        AND ((wFlowValid AND SHL(WORD#1, iBase)) <> WORD#0)
        AND ((wInputEnable AND SHL(WORD#1, i)) <> WORD#0)
        AND (rFlowLpm <= rSetpoint) THEN
        IF (wInputReaction AND SHL(WORD#1, i)) <> WORD#0 THEN
            axAbort[16 + i] := TRUE;
        ELSE
            axAlarm[16 + i] := TRUE;
        END_IF;
    END_IF;
END_FOR;

(* water pressure *)
rWaterBar := F_ReadFixed(awHolding[234], awHolding[235]);
IF ((wFlowValid AND WORD#16#0200) <> WORD#0)
    AND ((wInputEnable AND WORD#16#0040) <> WORD#0) THEN
    IF ((wInputReaction AND WORD#16#0040) <> WORD#0) AND (rWaterBar < C_WATER_ABORT_BAR) THEN
        axAbort[22] := TRUE;
    ELSIF rWaterBar < C_WATER_ALARM_BAR THEN
        axAlarm[22] := TRUE;
    END_IF;
END_IF;

(* compressed air pressure *)
rCdaBar := F_ReadFixed(awHolding[236], awHolding[237]);
IF ((wFlowValid AND WORD#16#0100) <> WORD#0)
    AND ((wInputEnable AND WORD#16#0100) <> WORD#0) THEN
    IF ((wInputReaction AND WORD#16#0100) <> WORD#0) AND (rCdaBar <= C_CDA_ABORT_BAR) THEN
        axAbort[23] := TRUE;
    ELSIF rCdaBar <= C_CDA_ALARM_BAR THEN
        axAlarm[23] := TRUE;
    END_IF;
END_IF;

(* chamber lid *)
IF ((wInputEnable AND WORD#16#0080) <> WORD#0) AND (NOT xLidClosed) THEN
    IF (wInputReaction AND WORD#16#0080) <> WORD#0 THEN
        axAbort[24] := TRUE;
    ELSE
        axAlarm[24] := TRUE;
    END_IF;
END_IF;

(* chamber pressure above 800 torr *)
IF arBandMeasured[0] > C_CHAMBER_MAX_TORR THEN
    axAlarm[25] := TRUE;
END_IF;

(* microwave generator faults while requested: only the microwave stops, latched until reset *)
IF xMwRequested THEN
    wMwTripNow := WORD#0;
    IF (wMwStatus AND WORD#16#8000) <> WORD#0 THEN wMwTripNow := wMwTripNow OR WORD#16#0001; END_IF;
    IF (wMwStatus AND WORD#16#2000) <> WORD#0 THEN wMwTripNow := wMwTripNow OR WORD#16#0002; END_IF;
    IF (wMwStatus AND WORD#16#4000) <> WORD#0 THEN wMwTripNow := wMwTripNow OR WORD#16#0004; END_IF;
    IF (wMwStatus AND WORD#16#1000) <> WORD#0 THEN wMwTripNow := wMwTripNow OR WORD#16#0008; END_IF;
    IF (wMwStatus AND WORD#16#0800) <> WORD#0 THEN wMwTripNow := wMwTripNow OR WORD#16#0010; END_IF;
    IF (wMwStatus AND WORD#16#0004) <> WORD#0 THEN wMwTripNow := wMwTripNow OR WORD#16#0020; END_IF;
    IF (wMwStatus AND WORD#16#0400) <> WORD#0 THEN wMwTripNow := wMwTripNow OR WORD#16#0040; END_IF;
    IF (wMwStatus AND WORD#16#0200) <> WORD#0 THEN wMwTripNow := wMwTripNow OR WORD#16#0080; END_IF;
    IF (wMwStatus AND WORD#16#0002) <> WORD#0 THEN wMwTripNow := wMwTripNow OR WORD#16#0200; END_IF;
    IF (wMwStatus AND WORD#16#0010) <> WORD#0 THEN axAlarm[40] := TRUE; END_IF;
    IF wMwTripNow <> WORD#0 THEN
        xMwTripActive := TRUE;
        wMwTripLatched := wMwTripLatched OR wMwTripNow;
    END_IF;
END_IF;

FOR i := 0 TO 9 DO
    IF (wMwTripLatched AND SHL(WORD#1, i)) <> WORD#0 THEN
        axAlarm[32 + i] := TRUE;
    END_IF;
END_FOR;

(* turbo pump faults *)
IF xTurboAnswering THEN
    IF (wTurboStatus AND WORD#16#0001) <> WORD#0 THEN axAlarm[48] := TRUE; END_IF;
    IF (wTurboStatus AND WORD#16#0002) <> WORD#0 THEN axAlarm[49] := TRUE; END_IF;
    IF (wTurboStatus AND WORD#16#0020) <> WORD#0 THEN axAlarm[50] := TRUE; END_IF;
    IF (wTurboStatus AND WORD#16#0040) <> WORD#0 THEN axAlarm[51] := TRUE; END_IF;
    IF (wTurboStatus AND WORD#16#0080) <> WORD#0 THEN axAlarm[52] := TRUE; END_IF;
    IF wTurboStatus = WORD#16#0108 THEN axAlarm[53] := TRUE; END_IF;
END_IF;

(* pack the flags into masks *)
FOR i := 0 TO 3 DO
    awAlarmMask[i] := WORD#0;
    awAbortMask[i] := WORD#0;
END_FOR;

xAnyAlarm := FALSE;
xAnyAbort := FALSE;

FOR i := 0 TO 63 DO
    iWord := i / 16;
    iBit := i MOD 16;
    IF axAlarm[i] THEN
        awAlarmMask[iWord] := awAlarmMask[iWord] OR SHL(WORD#1, iBit);
        xAnyAlarm := TRUE;
    END_IF;
    IF axAbort[i] THEN
        awAbortMask[iWord] := awAbortMask[iWord] OR SHL(WORD#1, iBit);
        xAnyAbort := TRUE;
    END_IF;
END_FOR;

(* abort: latches on its own, cleared by a reset from the hmi *)
xReset := xThresholdsOk AND ((awHolding[271] AND WORD#16#0002) <> WORD#0);

IF xAnyAbort AND (NOT xAbortActive) THEN
    xAbortActive := TRUE;
    uiAbortCount := uiAbortCount + UINT#1;
    FOR i := 0 TO 3 DO
        awAbortLatched[i] := awAbortMask[i];
    END_FOR;
END_IF;

(* on abort, inhibit everything that was on *)
IF xAbortActive THEN
    wGpvInhibit := wGpvInhibit OR awHolding[133];
    wVpvInhibit := wVpvInhibit OR awHolding[135];
    IF (awHolding[137] AND WORD#16#0002) <> WORD#0 THEN xForeVacInhibit := TRUE; END_IF;
    IF (awHolding[240] AND WORD#16#0001) <> WORD#0 THEN xTurboInhibit := TRUE; END_IF;
    IF (awHolding[192] AND WORD#16#0003) <> WORD#0 THEN xMwInhibit := TRUE; END_IF;
END_IF;

IF xMwTripActive AND ((awHolding[192] AND WORD#16#0003) <> WORD#0) THEN
    xMwInhibit := TRUE;
END_IF;

(* an inhibit clears once the hmi switches that output off *)
wGpvInhibit := wGpvInhibit AND awHolding[133];
wVpvInhibit := wVpvInhibit AND awHolding[135];
IF (awHolding[137] AND WORD#16#0002) = WORD#0 THEN xForeVacInhibit := FALSE; END_IF;
IF (awHolding[240] AND WORD#16#0001) = WORD#0 THEN xTurboInhibit := FALSE; END_IF;
IF (awHolding[192] AND WORD#16#0003) = WORD#0 THEN xMwInhibit := FALSE; END_IF;

(* reset from the hmi: microwave trip always, abort only when no cause is left *)
IF xReset AND (NOT xResetPrev) THEN
    xMwTripActive := FALSE;
    wMwTripLatched := WORD#0;
    IF NOT xAnyAbort THEN
        xAbortActive := FALSE;
        FOR i := 0 TO 3 DO
            awAbortLatched[i] := WORD#0;
        END_FOR;
    END_IF;
END_IF;
xResetPrev := xReset;

(* masks and status to the hmi *)
FOR i := 0 TO 3 DO
    awHolding[280 + i] := awAlarmMask[i];
    awHolding[284 + i] := awAbortMask[i];
    awHolding[288 + i] := awAbortLatched[i];
END_FOR;

wStatusWord := C_HMI_PROTOCOL;
IF xAbortActive THEN
    wStatusWord := wStatusWord OR WORD#16#0001;
END_IF;
IF xAnyAlarm THEN
    wStatusWord := wStatusWord OR WORD#16#0002;
END_IF;
IF xThresholdsOk THEN
    wStatusWord := wStatusWord OR WORD#16#0004;
END_IF;
IF xRetainWasBlank THEN
    wStatusWord := wStatusWord OR WORD#16#0008;
END_IF;
IF (wGpvInhibit <> WORD#0) OR (wVpvInhibit <> WORD#0)
    OR xForeVacInhibit OR xTurboInhibit OR xMwInhibit THEN
    wStatusWord := wStatusWord OR WORD#16#0010;
END_IF;
IF xMwTripActive THEN
    wStatusWord := wStatusWord OR WORD#16#0020;
END_IF;
awHolding[292] := wStatusWord;
awHolding[294] := wGpvInhibit;
awHolding[295] := wVpvInhibit;
awHolding[293] := UINT_TO_WORD(uiAbortCount);

(* ---- PRG_Cooling.st ---- *)
PROGRAM PRG_Cooling
(* cooling: water temperature and flow per circuit, water and air pressure *)
VAR CONSTANT
    (* scaling to volts and sensor units *)
    C_INT_TO_VOLT : REAL := 100.0;

    C_TEMP_ZERO  : REAL := 1.0;
    C_TEMP_SPAN  : REAL := 25.0;

    C_FLOW_ZERO  : REAL := 1.0;
    C_FLOW_SPAN  : REAL := 4.0;

    C_WATER_BAR_PER_VOLT : REAL := 1.666;
    C_CDA_BAR_PER_VOLT   : REAL := 1.0;

    (* circuit indices *)
    C_STAGE    : INT := 0;
    C_CHAMBER  : INT := 1;
    C_MWHEAD   : INT := 2;
    C_MWPOWER  : INT := 3;
    C_TUNER    : INT := 4;
    C_INTERNAL : INT := 5;
    C_EXTERNAL : INT := 6;

    C_CIRCUIT_MAX : INT := 6;

    (* module channels *)
    C_MOD2_BASE : INT := 8;
    C_WATER_CH  : INT := 14;
    C_CDA_CH    : INT := 15;

    (* flow channel of each circuit, temperature on the next one *)
    C_FLOW_CH : ARRAY[0..6] OF INT := [0, 2, 4, 6, 12, 8, 10];

    (* status bits for air and water pressure *)
    C_CDA_BIT   : INT := 8;
    C_WATER_BIT : INT := 9;
END_VAR
VAR
    i          : INT;
    iFlowCh    : INT;
    iTempCh    : INT;
    dwValue    : DWORD;
    wTempOk    : WORD;
    wFlowOk    : WORD;

    arChanVolt : ARRAY[0..15] OF REAL;
    axChanOk   : ARRAY[0..15] OF BOOL;

    arTempC    : ARRAY[0..6] OF REAL;
    arFlowLpm  : ARRAY[0..6] OF REAL;
    rWaterBar  : REAL;
    rCdaBar    : REAL;
END_VAR

(* both modules to volts, bad channels read as zero *)
FOR i := 0 TO 7 DO
    axChanOk[i] := (awCoolMod1Status[i] = WORD#16#0000);
    IF axChanOk[i] THEN
        arChanVolt[i] := INT_TO_REAL(WORD_TO_INT(awCoolMod1Value[i])) / C_INT_TO_VOLT;
    ELSE
        arChanVolt[i] := 0.0;
    END_IF;

    axChanOk[C_MOD2_BASE + i] := (awCoolMod2Status[i] = WORD#16#0000);
    IF axChanOk[C_MOD2_BASE + i] THEN
        arChanVolt[C_MOD2_BASE + i] := INT_TO_REAL(WORD_TO_INT(awCoolMod2Value[i])) / C_INT_TO_VOLT;
    ELSE
        arChanVolt[C_MOD2_BASE + i] := 0.0;
    END_IF;
END_FOR;

(* temperature and flow per circuit *)
wTempOk := WORD#0;
wFlowOk := WORD#0;
FOR i := 0 TO C_CIRCUIT_MAX DO
    iFlowCh := C_FLOW_CH[i];
    iTempCh := iFlowCh + 1;

    IF axChanOk[iTempCh] THEN
        wTempOk := wTempOk OR SHL(WORD#1, i);
    END_IF;
    IF axChanOk[iFlowCh] THEN
        wFlowOk := wFlowOk OR SHL(WORD#1, i);
    END_IF;

    IF arChanVolt[iTempCh] > C_TEMP_ZERO THEN
        arTempC[i] := (arChanVolt[iTempCh] - C_TEMP_ZERO) * C_TEMP_SPAN;
    ELSE
        arTempC[i] := 0.0;
    END_IF;

    IF arChanVolt[iFlowCh] > C_FLOW_ZERO THEN
        arFlowLpm[i] := (arChanVolt[iFlowCh] - C_FLOW_ZERO) * C_FLOW_SPAN;
    ELSE
        arFlowLpm[i] := 0.0;
    END_IF;
END_FOR;

(* compressed air and water pressure *)
rCdaBar := arChanVolt[C_CDA_CH] / C_CDA_BAR_PER_VOLT;
IF axChanOk[C_CDA_CH] THEN
    wFlowOk := wFlowOk OR SHL(WORD#1, C_CDA_BIT);
END_IF;

rWaterBar := arChanVolt[C_WATER_CH] / C_WATER_BAR_PER_VOLT;
IF axChanOk[C_WATER_CH] THEN
    wFlowOk := wFlowOk OR SHL(WORD#1, C_WATER_BIT);
END_IF;

(* everything to the hmi, registers 206..239 *)
FOR i := 0 TO C_CIRCUIT_MAX DO
    dwValue := F_ToFixed(arTempC[i]);
    awHolding[206 + 2*i] := DWORD_TO_WORD(dwValue);
    awHolding[207 + 2*i] := DWORD_TO_WORD(SHR(dwValue, 16));

    dwValue := F_ToFixed(arFlowLpm[i]);
    awHolding[220 + 2*i] := DWORD_TO_WORD(dwValue);
    awHolding[221 + 2*i] := DWORD_TO_WORD(SHR(dwValue, 16));
END_FOR;

dwValue := F_ToFixed(rWaterBar);
awHolding[234] := DWORD_TO_WORD(dwValue);
awHolding[235] := DWORD_TO_WORD(SHR(dwValue, 16));

dwValue := F_ToFixed(rCdaBar);
awHolding[236] := DWORD_TO_WORD(dwValue);
awHolding[237] := DWORD_TO_WORD(SHR(dwValue, 16));

awHolding[238] := wTempOk;
awHolding[239] := wFlowOk;

(* ---- PRG_Debug.st ---- *)
PROGRAM PRG_Debug
(* debug commands from the hmi system settings window *)
VAR
    wCommand     : WORD;
    wLastCommand : WORD;
    byCode       : BYTE;
    xFirstScan   : BOOL := TRUE;

    axMfcResetRequest : ARRAY[0..5] OF BOOL;
    afbMfcReset       : ARRAY[0..5] OF TP;
    xRebootRequest    : BOOL;
    fbRebootPulse     : TP;
    i : INT;
END_VAR
VAR CONSTANT
    C_RESET_ALL_MFC   : BYTE := 1;
    C_RESET_MFC_FIRST : BYTE := 2;
    C_REINIT_GAS      : BYTE := 20;
    C_REBOOT          : BYTE := 30;
END_VAR

(* register 148: low byte command, high byte sequence; run once per new word *)
wCommand := awHolding[148];
IF xFirstScan THEN
    wLastCommand := wCommand;
    xFirstScan := FALSE;
END_IF;

FOR i := 0 TO 5 DO
    axMfcResetRequest[i] := FALSE;
END_FOR;
xRebootRequest := FALSE;

IF wCommand <> wLastCommand THEN
    wLastCommand := wCommand;
    byCode := WORD_TO_BYTE(wCommand AND WORD#16#00FF);

    IF byCode = C_RESET_ALL_MFC THEN
        FOR i := 0 TO 5 DO
            axMfcResetRequest[i] := TRUE;
        END_FOR;
    ELSIF (byCode >= C_RESET_MFC_FIRST) AND (byCode <= C_RESET_MFC_FIRST + 5) THEN
        axMfcResetRequest[BYTE_TO_INT(byCode - C_RESET_MFC_FIRST)] := TRUE;
    ELSIF byCode = C_REINIT_GAS THEN
        uiDbgGasReinitCount := uiDbgGasReinitCount + 1;
    ELSIF byCode = C_REBOOT THEN
        xRebootRequest := TRUE;
    END_IF;
END_IF;

(* echo of the last accepted command *)
awHolding[149] := wLastCommand;

(* mfc link reset, 500 ms pulse per controller *)
FOR i := 0 TO 5 DO
    afbMfcReset[i](IN := axMfcResetRequest[i], PT := T#500MS);
END_FOR;
MFC_H2.xReset  := afbMfcReset[0].Q;
MFC_CH4.xReset := afbMfcReset[1].Q;
MFC_O2.xReset  := afbMfcReset[2].Q;
MFC_N2.xReset  := afbMfcReset[3].Q;
MFC_Ar.xReset  := afbMfcReset[4].Q;
MFC_H22.xReset := afbMfcReset[5].Q;

(* controller reboot: xDbgReboot is bound to the watchdog node reboot channel *)
fbRebootPulse(IN := xRebootRequest, PT := T#2S);
xDbgReboot := fbRebootPulse.Q;

(* ---- PRG_GasFlow.st ---- *)
PROGRAM PRG_GasFlow
(* mass flow controllers, six gas channels *)
VAR CONSTANT
    (* full scale per channel, sccm *)
    aFullScaleSccm : ARRAY[0..5] OF REAL := [1000.0, 100.0, 50.0, 1000.0, 10.0, 1000.0];
    C_INIT_DELAY_SCANS : INT := 3;
END_VAR
VAR
    xGasSubsystemEnable : BOOL;
    arSetpointSccm      : ARRAY[0..5] OF REAL;
    axSlaveError        : ARRAY[0..5] OF BOOL;
    aChState            : ARRAY[0..5] OF ST_GasChannelState;

    wGasStatus  : WORD;
    wChStatus   : WORD;
    dwValue     : DWORD;
    iBase       : INT;
    xAnyFault   : BOOL;
    xAllFault   : BOOL;
    rRaw        : REAL;
    iRawSetpoint: INT;
    i           : INT;
    uiReinitSeen: UINT;
END_VAR

(* gas enabled: hmi protocol ok, gas switched on, no abort *)
xGasSubsystemEnable := (awHolding[0] = WORD#1) AND ((awHolding[1] AND WORD#16#0008) <> WORD#0) AND (NOT xAbortActive);

(* link error per controller *)
axSlaveError[0] := MFC_H2.xError;
axSlaveError[1] := MFC_CH4.xError;
axSlaveError[2] := MFC_O2.xError;
axSlaveError[3] := MFC_N2.xError;
axSlaveError[4] := MFC_Ar.xError;
axSlaveError[5] := MFC_H22.xError;

(* setpoints from the hmi *)
FOR i := 0 TO 5 DO
    arSetpointSccm[i] := F_ReadFixed(awHolding[66 + i*5], awHolding[67 + i*5]);
END_FOR;

(* reinit request from the hmi debug window: regulating channels start init again *)
IF uiDbgGasReinitCount <> uiReinitSeen THEN
    uiReinitSeen := uiDbgGasReinitCount;
    FOR i := 0 TO 5 DO
        IF aChState[i].eInit = INIT_DONE THEN
            aChState[i].eInit := INIT_START;
        END_IF;
    END_FOR;
END_IF;

(* per channel: init, close, setpoint *)
FOR i := 0 TO 5 DO
    CASE aChState[i].eInit OF

        (* after enable, write ramp and mode one command at a time *)
        INIT_START:
            awRampTimeValue[i] := WORD#200;
            axRampTimeTrigger[i] := TRUE;
            aChState[i].iInitDelay := 0;
            aChState[i].eInit := INIT_RAMPTIME_HOLD;

        INIT_RAMPTIME_HOLD:
            axRampTimeTrigger[i] := FALSE;
            aChState[i].iInitDelay := aChState[i].iInitDelay + 1;
            IF aChState[i].iInitDelay >= C_INIT_DELAY_SCANS THEN
                awRampStepValue[i] := WORD#10;
                axRampStepTrigger[i] := TRUE;
                aChState[i].iInitDelay := 0;
                aChState[i].eInit := INIT_RAMPSTEP_HOLD;
            END_IF;

        INIT_RAMPSTEP_HOLD:
            axRampStepTrigger[i] := FALSE;
            aChState[i].iInitDelay := aChState[i].iInitDelay + 1;
            IF aChState[i].iInitDelay >= C_INIT_DELAY_SCANS THEN
                awRampEnValue[i] := WORD#1;
                axRampEnTrigger[i] := TRUE;
                aChState[i].iInitDelay := 0;
                aChState[i].eInit := INIT_RAMPEN_HOLD;
            END_IF;

        INIT_RAMPEN_HOLD:
            axRampEnTrigger[i] := FALSE;
            aChState[i].iInitDelay := aChState[i].iInitDelay + 1;
            IF aChState[i].iInitDelay >= C_INIT_DELAY_SCANS THEN
                awModeValue[i] := WORD#19;
                axModeTrigger[i] := TRUE;
                aChState[i].iInitDelay := 0;
                aChState[i].eInit := INIT_MODE_HOLD;
            END_IF;

        INIT_MODE_HOLD:
            axModeTrigger[i] := FALSE;
            aChState[i].iInitDelay := aChState[i].iInitDelay + 1;
            IF aChState[i].iInitDelay >= C_INIT_DELAY_SCANS THEN
                aChState[i].xRegulating := TRUE;
                aChState[i].xFaultActive := FALSE;
                aChState[i].xCloseConfirmed := FALSE;
                aChState[i].eInit := INIT_DONE;
            END_IF;

        (* regulating, close on disable or error *)
        INIT_DONE:
            IF (NOT xGasSubsystemEnable) OR axSlaveError[i] THEN
                aChState[i].xRegulating := FALSE;
                aChState[i].xFaultActive := xGasSubsystemEnable;
                awModeValue[i] := WORD#10;
                axModeTrigger[i] := TRUE;
                aChState[i].iInitDelay := 0;
                aChState[i].eInit := CLOSE_HOLD;
            END_IF;

        CLOSE_HOLD:
            axModeTrigger[i] := FALSE;
            aChState[i].iInitDelay := aChState[i].iInitDelay + 1;
            IF aChState[i].iInitDelay >= C_INIT_DELAY_SCANS THEN
                aChState[i].xCloseConfirmed := TRUE;
                aChState[i].eInit := CLOSED;
            END_IF;

        CLOSED:
            IF xGasSubsystemEnable AND (NOT axSlaveError[i]) THEN
                aChState[i].eInit := INIT_START;
            END_IF;

        ELSE
            aChState[i].eInit := INIT_START;
    END_CASE;

    (* setpoint to device units, sent only on change *)
    rRaw := arSetpointSccm[i] / aFullScaleSccm[i] * 10000.0;
    IF rRaw < 0.0 THEN
        rRaw := 0.0;
    END_IF;
    iRawSetpoint := REAL_TO_INT(rRaw + 0.5);
    IF iRawSetpoint > 10000 THEN
        iRawSetpoint := 10000;
    ELSIF iRawSetpoint < 0 THEN
        iRawSetpoint := 0;
    END_IF;

    IF iRawSetpoint <> aChState[i].iLastSetpointRaw THEN
        awSetpointRaw[i] := INT_TO_WORD(iRawSetpoint);
        axSetpointTrigger[i] := TRUE;
        aChState[i].iLastSetpointRaw := iRawSetpoint;
    ELSE
        axSetpointTrigger[i] := FALSE;
    END_IF;
END_FOR;

(* flow and status per channel to the hmi *)
xAnyFault := FALSE;
xAllFault := TRUE;
FOR i := 0 TO 5 DO
    iBase := 66 + i*5;

    dwValue := F_ToFixed(UINT_TO_REAL(WORD_TO_UINT(awMeasuredRaw[i])) / 10000.0 * aFullScaleSccm[i]);
    awHolding[iBase + 2] := DWORD_TO_WORD(dwValue);
    awHolding[iBase + 3] := DWORD_TO_WORD(SHR(dwValue, 16));

    wChStatus := WORD#0;
    IF aChState[i].xRegulating THEN
        wChStatus := wChStatus OR WORD#16#0001;
    END_IF;
    IF aChState[i].xFaultActive THEN
        wChStatus := wChStatus OR WORD#16#0002;
        xAnyFault := TRUE;
    ELSE
        xAllFault := FALSE;
    END_IF;
    IF aChState[i].xCloseConfirmed THEN
        wChStatus := wChStatus OR WORD#16#0004;
    END_IF;
    IF (NOT xGasSubsystemEnable) AND (NOT aChState[i].xFaultActive) THEN
        wChStatus := wChStatus OR WORD#16#0008;
    END_IF;
    awHolding[iBase + 4] := wChStatus;
END_FOR;

(* overall gas status *)
wGasStatus := WORD#0;
IF NOT xAllFault THEN
    wGasStatus := wGasStatus OR WORD#16#0001;
END_IF;
IF xAnyFault THEN
    wGasStatus := wGasStatus OR WORD#16#0002;
END_IF;
IF xAllFault THEN
    wGasStatus := wGasStatus OR WORD#16#0004;
END_IF;
IF xGasSubsystemEnable THEN
    wGasStatus := wGasStatus OR WORD#16#0008;
END_IF;
awHolding[64] := wGasStatus;
awHolding[65] := awHolding[65] + WORD#1;

(* link errors per channel, debug for the first two channels *)
wChStatus := WORD#0;
FOR i := 0 TO 5 DO
    IF axSlaveError[i] THEN
        wChStatus := wChStatus OR SHL(WORD#1, i);
    END_IF;
END_FOR;
awHolding[96] := wChStatus;
awHolding[97] := awMeasuredRaw[0];
CASE aChState[0].eInit OF
    INIT_START:         awHolding[98] := WORD#0;
    INIT_RAMPTIME_HOLD: awHolding[98] := WORD#1;
    INIT_RAMPSTEP_HOLD: awHolding[98] := WORD#2;
    INIT_RAMPEN_HOLD:   awHolding[98] := WORD#3;
    INIT_MODE_HOLD:     awHolding[98] := WORD#4;
    INIT_DONE:          awHolding[98] := WORD#5;
    CLOSE_HOLD:         awHolding[98] := WORD#6;
    CLOSED:             awHolding[98] := WORD#7;
END_CASE;

CASE aChState[1].eInit OF
    INIT_START:         awHolding[99] := WORD#0;
    INIT_RAMPTIME_HOLD: awHolding[99] := WORD#1;
    INIT_RAMPSTEP_HOLD: awHolding[99] := WORD#2;
    INIT_RAMPEN_HOLD:   awHolding[99] := WORD#3;
    INIT_MODE_HOLD:     awHolding[99] := WORD#4;
    INIT_DONE:          awHolding[99] := WORD#5;
    CLOSE_HOLD:         awHolding[99] := WORD#6;
    CLOSED:             awHolding[99] := WORD#7;
END_CASE;

(* ---- PRG_GasValves.st ---- *)
PROGRAM PRG_GasValves
(* gas valves gpv1..gpv8 *)
VAR
    wGpvCommand : WORD;
    wGpvStatus  : WORD;
    i : INT;
END_VAR

(* command from the hmi, all closed on abort *)
IF xAbortActive THEN
    wGpvCommand := WORD#0;
ELSE
    wGpvCommand := awHolding[133] AND (NOT wGpvInhibit);
END_IF;

(* to the outputs *)
FOR i := 1 TO 8 DO
    axGpvOutput[i] := (wGpvCommand AND SHL(WORD#1, i - 1)) <> WORD#0;
END_FOR;

(* actual output state back to the hmi *)
wGpvStatus := WORD#0;
FOR i := 1 TO 8 DO
    IF axGpvOutput[i] THEN
        wGpvStatus := wGpvStatus OR SHL(WORD#1, i - 1);
    END_IF;
END_FOR;

awHolding[134] := wGpvStatus;

(* ---- PRG_Pyrometers.st ---- *)
PROGRAM PRG_Pyrometers
(* pyrometers *)
VAR
    uPyroValue : U_DWORD_REAL;

    rPyroRxtCh1     : REAL;
    rPyroRxtCh2     : REAL;
    rPyroRxtRatio   : REAL;
    wPyroRxtStatus  : WORD;

    dwValue : DWORD;

    fbCommOk       : TON;
    fbConfirmPulse : TP;
    xPyroReconnectRequest : BOOL;
END_VAR

(* link ok after 4 s without errors *)
fbCommOk(IN := NOT PYRO_RXT.xError, PT := T#4S);

(* reconnect request from the hmi, register 170 bit 0 *)
xPyroReconnectRequest := (awHolding[170] AND WORD#16#0001) <> WORD#0;

(* rxt pyrometer: ch1, ch2 and ratio *)
uPyroValue.dwValue := SHL(WORD_TO_DWORD(awPyroRxtCh1Raw[1]), 16) OR WORD_TO_DWORD(awPyroRxtCh1Raw[0]);
rPyroRxtCh1 := uPyroValue.rValue;
uPyroValue.dwValue := SHL(WORD_TO_DWORD(awPyroRxtCh2Raw[1]), 16) OR WORD_TO_DWORD(awPyroRxtCh2Raw[0]);
rPyroRxtCh2 := uPyroValue.rValue;
uPyroValue.dwValue := SHL(WORD_TO_DWORD(awPyroRxtRatioRaw[1]), 16) OR WORD_TO_DWORD(awPyroRxtRatioRaw[0]);
rPyroRxtRatio := uPyroValue.rValue;

(* temperatures to the hmi, registers 160..165 *)
dwValue := F_ToFixed(rPyroRxtCh1);
awHolding[160] := DWORD_TO_WORD(dwValue);
awHolding[161] := DWORD_TO_WORD(SHR(dwValue, 16));
dwValue := F_ToFixed(rPyroRxtCh2);
awHolding[162] := DWORD_TO_WORD(dwValue);
awHolding[163] := DWORD_TO_WORD(SHR(dwValue, 16));
dwValue := F_ToFixed(rPyroRxtRatio);
awHolding[164] := DWORD_TO_WORD(dwValue);
awHolding[165] := DWORD_TO_WORD(SHR(dwValue, 16));

(* status: link and channel overload *)
wPyroRxtStatus := WORD#0;
IF fbCommOk.Q THEN
    wPyroRxtStatus := wPyroRxtStatus OR WORD#16#0001;
END_IF;
IF (wPyroRxtAdcStatus AND WORD#16#0001) <> WORD#0 THEN
    wPyroRxtStatus := wPyroRxtStatus OR WORD#16#0002;
END_IF;
IF (wPyroRxtAdcStatus AND WORD#16#0002) <> WORD#0 THEN
    wPyroRxtStatus := wPyroRxtStatus OR WORD#16#0004;
END_IF;
IF NOT fbCommOk.Q THEN
    wPyroRxtStatus := wPyroRxtStatus OR WORD#16#0008;
END_IF;
awHolding[166] := wPyroRxtStatus;
awHolding[167] := wPyroRxtDevStatus;

(* reconnect to the pyrometer after a link error *)
fbConfirmPulse(IN := xPyroReconnectRequest, PT := T#500MS);
PYRO_RXT.xConfirmError := fbConfirmPulse.Q;

(* ---- PRG_Thyracont.st ---- *)
PROGRAM PRG_Thyracont
(* thyracont vacuum gauge *)
VAR
    fbThyracont : FB_ThyracontAscii;
    udiThyracontPort : UDINT := 5;
    udiThyracontAddress : UDINT := 1;
    uValue : U_DWORD_REAL;

END_VAR

(* poll the gauge *)
fbThyracont(
    xEnable := TRUE,
    udiPort := udiThyracontPort,
    udiAddress := udiThyracontAddress,
    udiBaudrate := 9600,
    tPollInterval := T#0MS);

(* pressure and status to the hmi, registers 140..147 *)
uValue.rValue := fbThyracont.rPressureTorr;
awHolding[140] := DWORD_TO_WORD(uValue.dwValue);
awHolding[141] := DWORD_TO_WORD(SHR(uValue.dwValue, 16));
uValue.rValue := fbThyracont.rPressureMbar;
awHolding[142] := DWORD_TO_WORD(uValue.dwValue);
awHolding[143] := DWORD_TO_WORD(SHR(uValue.dwValue, 16));
awHolding[144] := fbThyracont.wStatusFlags;
awHolding[145] := fbThyracont.wErrorCode;
awHolding[146] := DWORD_TO_WORD(fbThyracont.udiCycle);
awHolding[147] := DWORD_TO_WORD(SHR(fbThyracont.udiCycle, 16));

(* ---- PRG_TurboPump.st ---- *)
PROGRAM PRG_TurboPump
(* turbo pump *)
VAR
    xCommandValid    : BOOL;
    xRunRequest      : BOOL;
    wCommandWanted   : WORD;
    wCommandSent     : WORD;
    xCommandIssued   : BOOL;

    wLatchedStatus : WORD;
    wLinkStatus    : WORD;
END_VAR
VAR CONSTANT
    C_CMD_RUN  : WORD := WORD#16#0008;
    C_CMD_STOP : WORD := WORD#16#0003;
END_VAR

(* command from the hmi, stop only on abort *)
xCommandValid := ((awHolding[240] AND WORD#16#8000) <> WORD#0) OR xAbortActive;
xRunRequest := ((awHolding[240] AND WORD#16#0001) <> WORD#0) AND (NOT xAbortActive) AND (NOT xTurboInhibit);

IF xRunRequest THEN
    wCommandWanted := C_CMD_RUN;
ELSE
    wCommandWanted := C_CMD_STOP;
END_IF;

(* send to the drive only when the command changes *)
IF xCommandValid AND ((NOT xCommandIssued) OR (wCommandWanted <> wCommandSent)) THEN
    wTurboCommandValue := wCommandWanted;
    xTurboCommandTrigger := TRUE;
    wCommandSent := wCommandWanted;
    xCommandIssued := TRUE;
ELSE
    xTurboCommandTrigger := FALSE;
END_IF;

(* status to the hmi *)
wLatchedStatus := WORD#0;
IF wCommandSent = C_CMD_RUN THEN
    wLatchedStatus := wLatchedStatus OR WORD#16#0001;
END_IF;
IF xCommandIssued THEN
    wLatchedStatus := wLatchedStatus OR WORD#16#0002;
END_IF;

wLinkStatus := WORD#0;
IF NOT TURBO_PUMP.xError THEN
    wLinkStatus := wLinkStatus OR WORD#16#0001;
END_IF;

awHolding[241] := wLatchedStatus;
awHolding[242] := awTurboStatusRaw[0];
awHolding[243] := awTurboStatusRaw[1];
awHolding[244] := awTurboStatusRaw[2];
awHolding[245] := awTurboStatusRaw[3];
awHolding[246] := wTurboTempRaw AND WORD#16#00FF;
awHolding[247] := wLinkStatus;

(* ---- PRG_VacuumOutputs.st ---- *)
PROGRAM PRG_VacuumOutputs
(* vacuum valves and pumps *)
VAR
    wVpvCommand  : WORD;
    wVpvStatus   : WORD;
    wPumpCommand : WORD;
    wPumpStatus  : WORD;
    i : INT;
END_VAR

(* valves: command from the hmi, all closed on abort *)
IF xAbortActive THEN
    wVpvCommand := WORD#0;
ELSE
    wVpvCommand := awHolding[135] AND (NOT wVpvInhibit);
END_IF;

FOR i := 1 TO 8 DO
    axVpvOutput[i] := (wVpvCommand AND SHL(WORD#1, i - 1)) <> WORD#0;
END_FOR;

(* valve state to the hmi *)
wVpvStatus := WORD#0;
FOR i := 1 TO 8 DO
    IF axVpvOutput[i] THEN
        wVpvStatus := wVpvStatus OR SHL(WORD#1, i - 1);
    END_IF;
END_FOR;

awHolding[136] := wVpvStatus;

(* water pump and forevacuum pump, forevacuum off on abort *)
wPumpCommand := awHolding[137];
xWaterPumpOutput := (wPumpCommand AND WORD#16#0001) <> WORD#0;
xForeVacPumpOutput := ((wPumpCommand AND WORD#16#0002) <> WORD#0) AND (NOT xAbortActive) AND (NOT xForeVacInhibit);

(* pump state to the hmi *)
wPumpStatus := WORD#0;
IF xWaterPumpOutput THEN
    wPumpStatus := wPumpStatus OR WORD#16#0001;
END_IF;
IF xForeVacPumpOutput THEN
    wPumpStatus := wPumpStatus OR WORD#16#0002;
END_IF;

awHolding[138] := wPumpStatus;
